(* IEC 61131-3 sources: Codesys-Github-Test/project-view/Controller_1/Plc Logic/Application, 2 files *)

(* ---- Motion_PRG.st ---- *)
PROGRAM Motion_PRG
VAR
END_VAR
END_PROGRAM

(* ---- PLC_PRG.st ---- *)
PROGRAM PLC_PRG
VAR
	i:INT;
	j:INT;
	test:INT;
END_VAR
// --- implementation ---
i:=i+1;
j:=j+1;
test:=i+j;

//FK趙公測試
//20261019翔帥修改
//翔帥測試1020
//123456再次測試
//5678丹青媽媽
////趙公工小鳥鳥
//翔大雕VS小鳥鳥
//第三次測試123
//翔大雕第四次測試
END_PROGRAM
